// SIMATIC S7-200 project (STEP 7-Micro/WIN), CPU 226 CN REL 02.01

SYMBOL_TABLE USUARIO1
SI1              I0.0     // Sensor de riel
FCI              I0.1     // Final de carrera derecha
FCF              I0.2     // Final de carrera izquierda
QS               I2.4     // Pulsador de parada
SB_1             I2.5     // Pulsador de marcha
SB_2             I2.6     // Zeta de emergencia
SA               I2.7     // Selector de modo
PULSO            Q0.0     // Pulso
DIR              Q0.1     // Direccion
                 Q0.3     // Cilndro neumatico vertical
                 Q0.4     // Cilindro rotarorio anti horario
                 Q0.5     // Cilindro rotatorio horario
                 Q0.6     // Cilindro horizontal
                 Q0.7     // Garra cerrada
                 Q1.0     // Garra abierta
HL1              Q1.5     // Piloto Amarillo
HL2              Q1.6     // Piloto Verde
HL3              Q1.7     // Piloto Rojo
END_SYMBOL_TABLE

ORGANIZATION_BLOCK PRINCIPAL:OB1
TITLE=COMENTARIOS DEL PROGRAMA
BEGIN
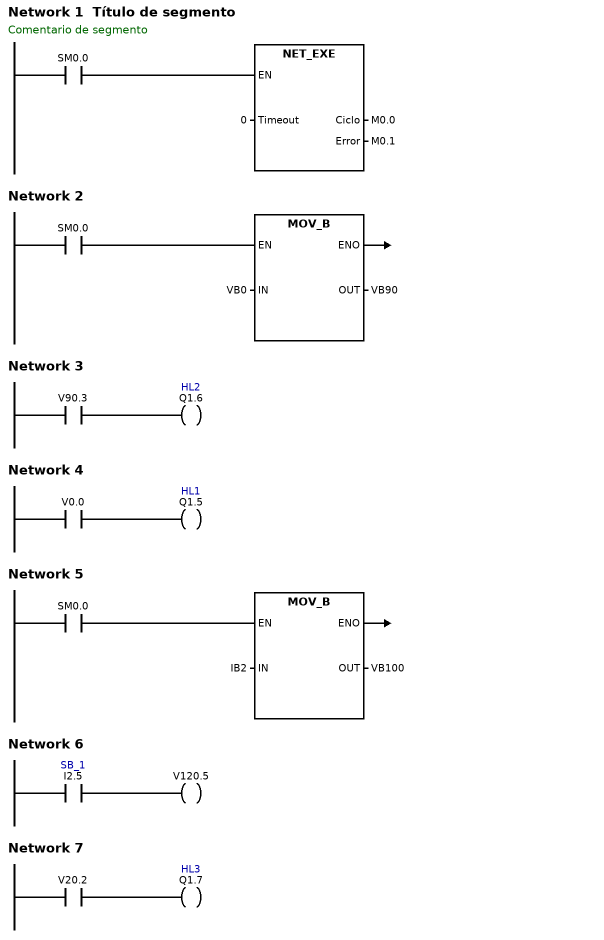
Network 1 // Título de segmento
// Comentario de segmento
LD     SM0.0
CALL   NET_EXE:SBR1, 0, M0.0, M0.1
Network 2
LD     SM0.0
MOVB   VB0, VB90
Network 3
LD     V90.3
=      HL2:Q1.6
Network 4
LD     V0.0
=      HL1:Q1.5
Network 5
LD     SM0.0
MOVB   IB2, VB100
Network 6
LD     SB_1:I2.5
=      V120.5
Network 7
LD     V20.2
=      HL3:Q1.7
END_ORGANIZATION_BLOCK

// SBR1: protected block, not included
